// TIA Portal V20 export
Screen "Hemming Process"  395x350
  ScreenItem "Robot Name" at 2,2 size 393x48  Type=HmiIOField
  ScreenItem "Background" at -24,46 size 419x300  Type=HmiRectangle
  ScreenItem "Cancel Mode" at 315,4 size 76x42  Type=HmiButton
  ScreenItem "矩形_4" at 31,99 size 324x76  Type=HmiRectangle
  ScreenItem "Text Field In Auto On_9" at 34,101 size 318x21  Type=HmiTextBox
  ScreenItem "Text Field Home Position_17" at 34,124 size 318x21  Type=HmiTextBox
  ScreenItem "Text field Robot Status_5" at 33,70 size 324x26  Type=HmiTextBox
  ScreenItem "Text Field System Ready_9" at 34,148 size 318x21  Type=HmiTextBox
